(* Logix 5000 project; controller R400_500_XLS vendor 1 type 14 code 216 rev 31.11; software revision 31.01; part 4 of 32 *)
(* tags used below, declared in another part *)
   Alarm : SINT;   // Wait 3 seconds
   bResetAllCycle : BOOL;
   ClearIndex : DINT;
   Condenser : INT;
   Cycles : UDT_CYCLE[11];
   FINAL_RINSE_MAX_NBR : INT;   // Maximum nimber of final rinse
   LowPressAlmSp : REAL;   // Pump pressure too low setpoint
   MaxTrtTempSp : REAL;
   PrintoutMSGTranslation : DINT;   // Grapcet for Printout Message Translation
   PrintoutMSGTranslationONS : INT;
   PURE_WATER_HEATING_TIME : DINT;   // Time before an alarm is thrown when the pure water tank is heating
   PWTnkTempAlmSp : REAL;   // Pure water tank temperature too high setpoint
   String : STRING[50];   // String
   SumpTempAlmSp : REAL;   // Sump temperature too high setpoint
   tHandshakeToggle : TIMER;
   Tmr : TIMER[107];
   bFactoryReset : BOOL;
   bFactoryResetCompleted : BOOL;
   BoilingValue : REAL;
   bONSFactoryReset : BOOL;
   bResetHardwareOptions : BOOL;
   bResetModulesConfiguration : BOOL;
   bResetSystemOptions : BOOL;
   Cfg_10_Modules : BOOL;   // Chassis is configured 10 slots
   Cfg_11_Modules : BOOL;
   ChangeLanguage : BOOL;   // Tag Changed By HMI To Start Printout Message Translation
   COOLING_PHASE_TIME : DINT;   // Time of the cooling phase when time based drying
   CycleCounter : DINT;
   DrainExtensionTime : DINT;
   EmailSMSInt : INT[8];   // Email & SMS Notification Integer
   FC45_NbCycBeforeMaint : DINT;
   I_Chem_Cond : DINT;   // Chemical water conductivity
   I_Chm_1_Lvl_Sw : BOOL;   // Chemical Pump #1 level switch
   I_Chm_2_Lvl_Sw : BOOL;   // Chemical Pump #2 level switch
   I_Chm_3_Lvl_Sw : BOOL;   // Chemical Pump #3 level switch
   I_Chm_4_Lvl_Sw : BOOL;   // Chemical Pump #4 level switch
   I_Dry_RTD : DINT;   // Drying RTD
   I_Final_Rinse_Cond : DINT;   // Final rinse water conductivity
   I_Ld_Dr_Cls_Sw : BOOL;   // Load door close
   I_Ld_Dr_Obs_Sw : BOOL;   // Load door obstruction switch
   I_MCR : BOOL;   // MCR input
   I_Mtr_Ovrld : BOOL;   // Motor overload
   I_Pump_Press : DINT;   // Recirculation pump pressure
   I_Pure_Water_Filling_Auth : BOOL;
   I_Pw_Tnk_Lvl_Sw : BOOL;   // Pure water tank level switch
   I_Pw_Tnk_RTD : DINT;   // Pure water tank RTD
   I_Pw_Tnk_Sft_Lvl_Sw : BOOL;   // Pure water tank safety level switch
   I_Shlf_Sw : BOOL;   // Shelf switch
   I_Smp_Lvl_Hgh : BOOL;   // Sump high level switch
   I_Smp_Lvl_Lw : BOOL;   // Sump low level switch
   I_Smp_RTD : DINT;   // Sump RTD
   I_Smp_Sft_Lvl_Sw : BOOL;   // Sump safety level switch
   I_Unld_Dr_Cls_Sw : BOOL;   // Unload door close
   I_Unld_Dr_Obs_Sw : BOOL;   // Unload door obstruction switch
   I_UnldDr_ClseSlnce_Bttn : BOOL;   // Door Close/ Silence button Unload Side
   I_UnldDr_Opn_Bttn : BOOL;   // Door Open button Unload side
   iDelayBeforeFillingAuthAlarmMM : DINT;
   iDelayBeforeFillingAuthAlarmSS : DINT;
   iInactivityLogoutTime : DINT;   // Inactivity Logout Time In Minutes
   iPWClosingDelayMM : DINT;
   iPWClosingDelaySS : DINT;
   msg : BOOL[512];
   MsgIterator : DINT;   // Iterator to Iterate Through all Printout Mesage
   MsgNumbers : DINT;
   NOT_USED : SINT[3];
   NumInput : UDT_NUMERIC_INPUT[65];   // Numeric input
   NumInputReal : UDT_NUMERIC_INPUT_REAL[17];
   PrintoutMsgHandshake : BOOL;   // Flag Send to HMI to Acknowledge Reception of Message
   PrintoutMsgNotification : BOOL[512];   // Flag Send by HMI when a Message is sended to PLC
   Screen_Ctrl : DINT;   // PLC Screen Request
   SumpAlarmFillTime : DINT;
   Tpb : DINT[11];
   Unit : Hrdwre;   // Unit Configuration
(* MainProgram, continued *)

ROUTINE EMAIL_SEND   (* ladder *)
// SEND EMAIL
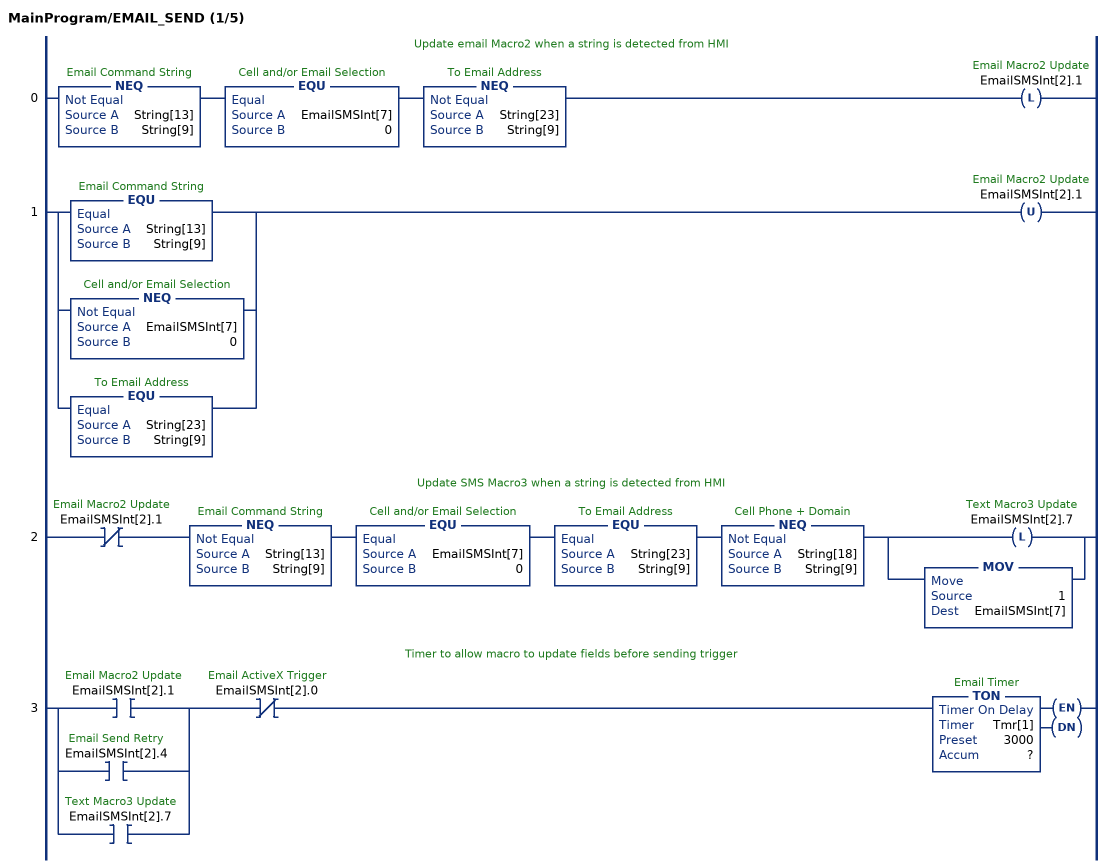
   // Update email Macro2 when a string is detected from HMI
   0: NEQ(String[13],String[9])EQU(EmailSMSInt[7],0)NEQ(String[23],String[9])OTL(EmailSMSInt[2].1);
   1: [EQU(String[13],String[9]) ,NEQ(EmailSMSInt[7],0) ,EQU(String[23],String[9]) ]OTU(EmailSMSInt[2].1);
   // Update SMS Macro3 when a string is detected from HMI
   2: XIO(EmailSMSInt[2].1)NEQ(String[13],String[9])EQU(EmailSMSInt[7],0)EQU(String[23],String[9])NEQ(String[18],String[9])[OTL(EmailSMSInt[2].7) ,MOV(1,EmailSMSInt[7]) ];
   // Timer to allow macro to update fields before sending trigger
   3: [XIC(EmailSMSInt[2].1) ,XIC(EmailSMSInt[2].4) ,XIC(EmailSMSInt[2].7) ]XIO(EmailSMSInt[2].0)TON(Tmr[1],?,?);
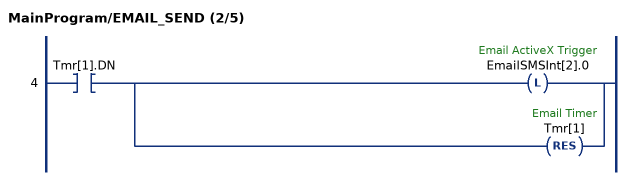
   4: XIC(Tmr[1].DN)[OTL(EmailSMSInt[2].0) ,RES(Tmr[1]) ];
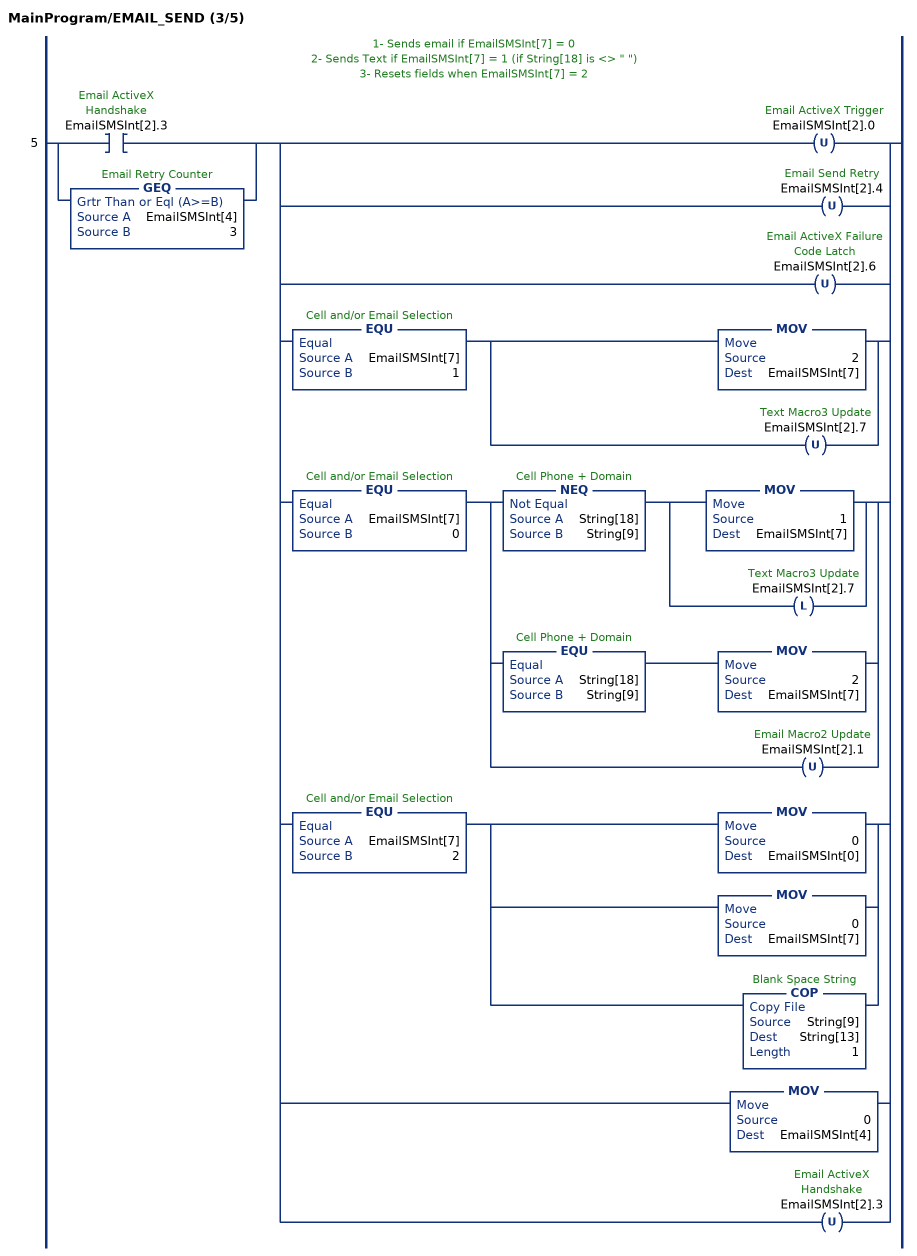
   // 1- Sends email if EmailSMSInt[7] = 0
   // 2- Sends Text if EmailSMSInt[7] = 1 (if String[18] is <> " ")
   // 3- Resets fields when EmailSMSInt[7] = 2
   5: [XIC(EmailSMSInt[2].3) ,GEQ(EmailSMSInt[4],3) ][OTU(EmailSMSInt[2].0) ,OTU(EmailSMSInt[2].4) ,OTU(EmailSMSInt[2].6) ,EQU(EmailSMSInt[7],1) [MOV(2,EmailSMSInt[7]) ,OTU(EmailSMSInt[2].7) ] ,EQU(EmailSMSInt[7],0) [NEQ(String[18],String[9]) [MOV(1,EmailSMSInt[7]) ,OTL(EmailSMSInt[2].7) ] ,EQU(String[18],String[9]) MOV(2,EmailSMSInt[7]) ,OTU(EmailSMSInt[2].1) ] ,EQU(EmailSMSInt[7],2) [MOV(0,EmailSMSInt[0]) ,MOV(0,EmailSMSInt[7]) ,COP(String[9],String[13],1) ] ,MOV(0,EmailSMSInt[4]) ,OTU(EmailSMSInt[2].3) ];
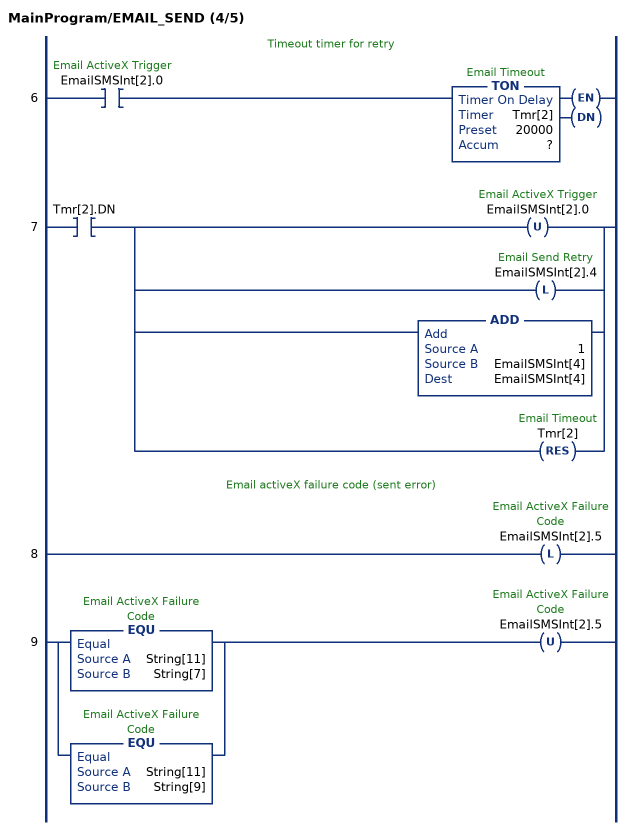
   // Timeout timer for retry
   6: XIC(EmailSMSInt[2].0)TON(Tmr[2],?,?);
   7: XIC(Tmr[2].DN)[OTU(EmailSMSInt[2].0) ,OTL(EmailSMSInt[2].4) ,ADD(1,EmailSMSInt[4],EmailSMSInt[4]) ,RES(Tmr[2]) ];
   // Email activeX failure code (sent error)
   8: OTL(EmailSMSInt[2].5);
   9: [EQU(String[11],String[7]) ,EQU(String[11],String[9]) ]OTU(EmailSMSInt[2].5);
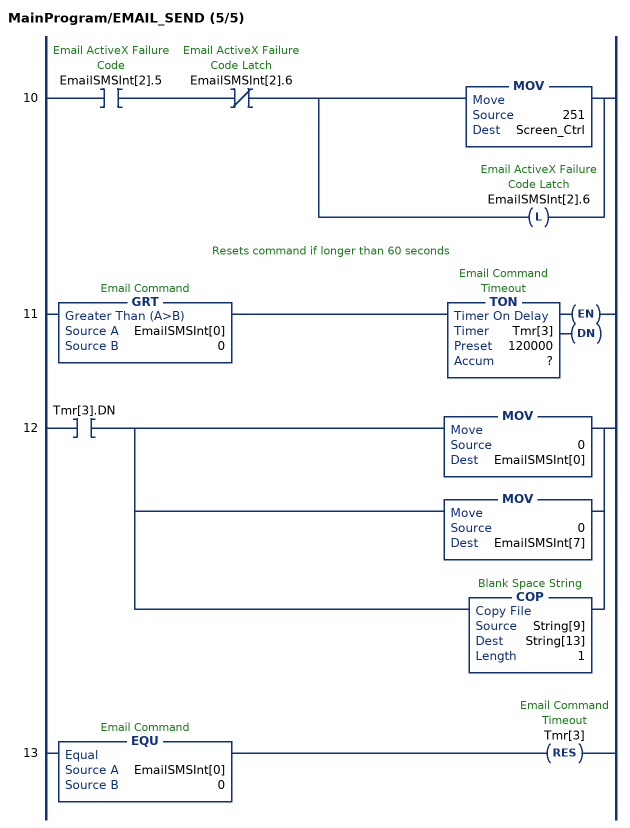
   10: XIC(EmailSMSInt[2].5)XIO(EmailSMSInt[2].6)[MOV(251,Screen_Ctrl) ,OTL(EmailSMSInt[2].6) ];
   // Resets command if longer than 60 seconds
   11: GRT(EmailSMSInt[0],0)TON(Tmr[3],?,?);
   12: XIC(Tmr[3].DN)[MOV(0,EmailSMSInt[0]) ,MOV(0,EmailSMSInt[7]) ,COP(String[9],String[13],1) ];
   13: EQU(EmailSMSInt[0],0)RES(Tmr[3]);
END_ROUTINE

ROUTINE FactoryReset   (* ladder *)
// This Routine contains logic to manage the Factory Reset
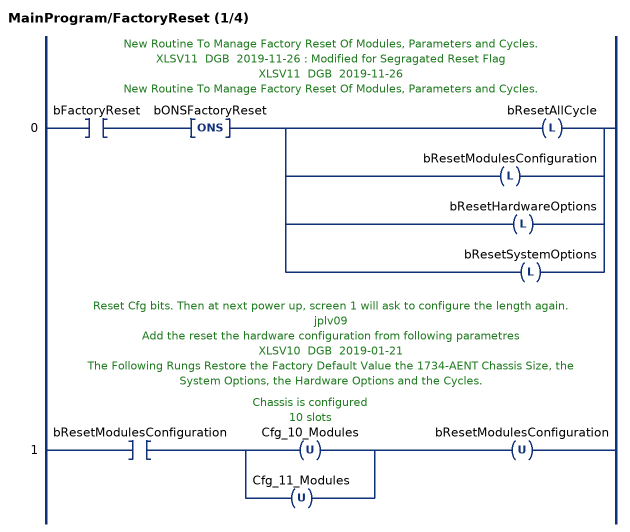
   // New Routine To Manage Factory Reset Of Modules, Parameters and Cycles.
   // XLSV11  DGB  2019-11-26 : Modified for Segragated Reset Flag
   // XLSV11  DGB  2019-11-26
   // New Routine To Manage Factory Reset Of Modules, Parameters and Cycles.
   0: XIC(bFactoryReset)ONS(bONSFactoryReset)[OTL(bResetAllCycle) ,OTL(bResetModulesConfiguration) ,OTL(bResetHardwareOptions) ,OTL(bResetSystemOptions) ];
   // Reset Cfg bits. Then at next power up, screen 1 will ask to configure the length again.
   // jplv09
   // Add the reset the hardware configuration from following parametres
   // XLSV10  DGB  2019-01-21
   // The Following Rungs Restore the Factory Default Value the 1734-AENT Chassis Size, the System Options, the Hardware Options and the Cycles.
   1: XIC(bResetModulesConfiguration)[OTU(Cfg_10_Modules) ,OTU(Cfg_11_Modules) ]OTU(bResetModulesConfiguration);
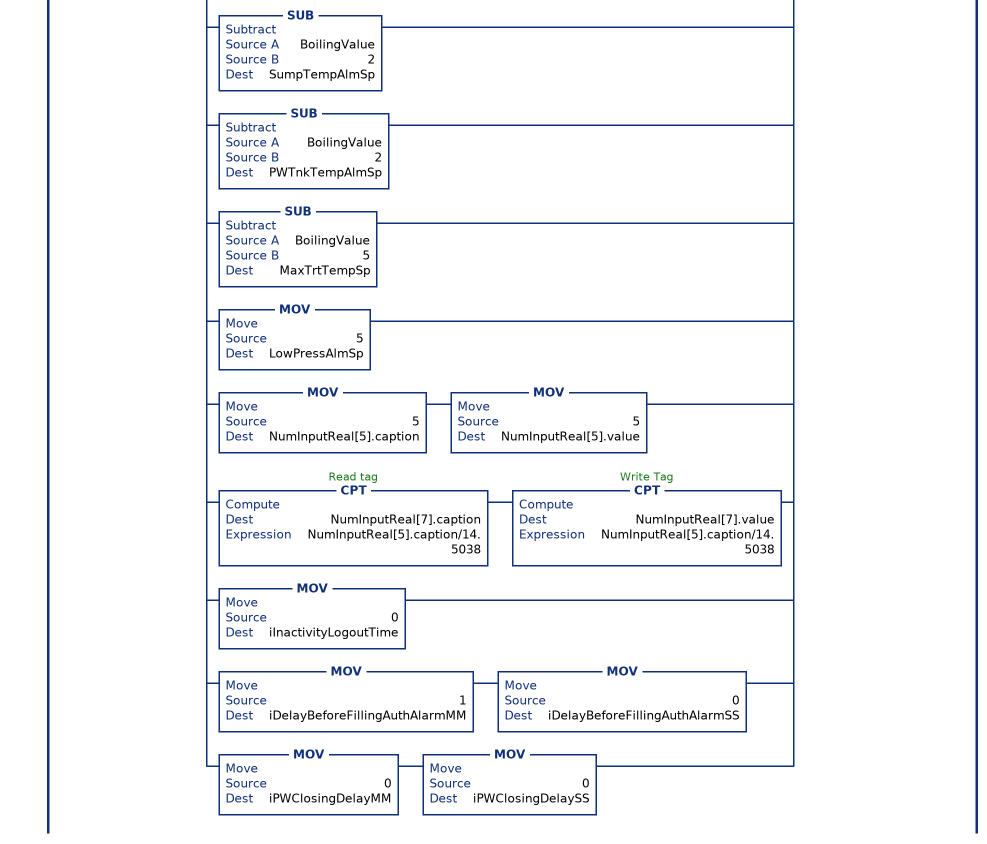
   // XLSV10  DGB  2019-01-21
   // New Rung to Restore the Factory Default Value of System Options
   // XLSV13  DGB  2021-03-16 : PW Filling Handshake : Added Pure Water Closing Delay & Delay Before Fill Auth Alarm Message
   2: XIC(bResetSystemOptions)[MOV(0,CycleCounter) ,MOV(1000,FC45_NbCycBeforeMaint) ,[MOV(120000,SumpAlarmFillTime) ,MOV(2,NumInput[9].caption) MOV(2,NumInput[9].value) ,MOV(0,NumInput[10].caption) MOV(0,NumInput[10].value) ] ,[MOV(20000,Tmr[88].PRE) ,MOV(20,NumInput[52].caption) MOV(20,NumInput[52].value) ] ,[MOV(480000,Tmr[37].PRE) ,MOV(8,NumInput[38].caption) MOV(8,NumInput[38].value) ,MOV(0,NumInput[39].caption) MOV(0,NumInput[39].value) ] ,[MOV(1200000,PURE_WATER_HEATING_TIME) ,MOV(20,NumInput[40].caption) MOV(20,NumInput[40].value) ,MOV(0,NumInput[41].caption) MOV(0,NumInput[41].value) ] ,[MOV(9,FINAL_RINSE_MAX_NBR) ,MOV(9,NumInput[42].caption) MOV(9,NumInput[42].value) ] ,[MOV(0,DrainExtensionTime) ,MOV(0,NumInput[43].caption) MOV(0,NumInput[43].value) ] ,[MOV(120000,Tmr[31].PRE) ,MOV(2,NumInput[44].caption) MOV(2,NumInput[44].value) ,MOV(0,NumInput[45].caption) MOV(0,NumInput[45].value) ] ,[MOV(120000,COOLING_PHASE_TIME) ,MOV(2,NumInput[47].caption) MOV(2,NumInput[47].value) ,MOV(0,NumInput[48].caption) MOV(0,NumInput[48].value) ] ,[MOV(0,NumInput[46].caption) MOV(0,NumInput[46].value) ,CPT(BoilingValue,100.03) ,SUB(BoilingValue,2,SumpTempAlmSp) ,SUB(BoilingValue,2,PWTnkTempAlmSp) ,SUB(BoilingValue,5,MaxTrtTempSp) ] ,[MOV(5,LowPressAlmSp) ,MOV(5,NumInputReal[5].caption) MOV(5,NumInputReal[5].value) ,CPT(NumInputReal[7].caption,NumInputReal[5].caption/14.5038) CPT(NumInputReal[7].value,NumInputReal[5].caption/14.5038) ] ,MOV(0,iInactivityLogoutTime) ,MOV(1,iDelayBeforeFillingAuthAlarmMM) MOV(0,iDelayBeforeFillingAuthAlarmSS) ,MOV(0,iPWClosingDelayMM) MOV(0,iPWClosingDelaySS) ]OTU(bResetSystemOptions);
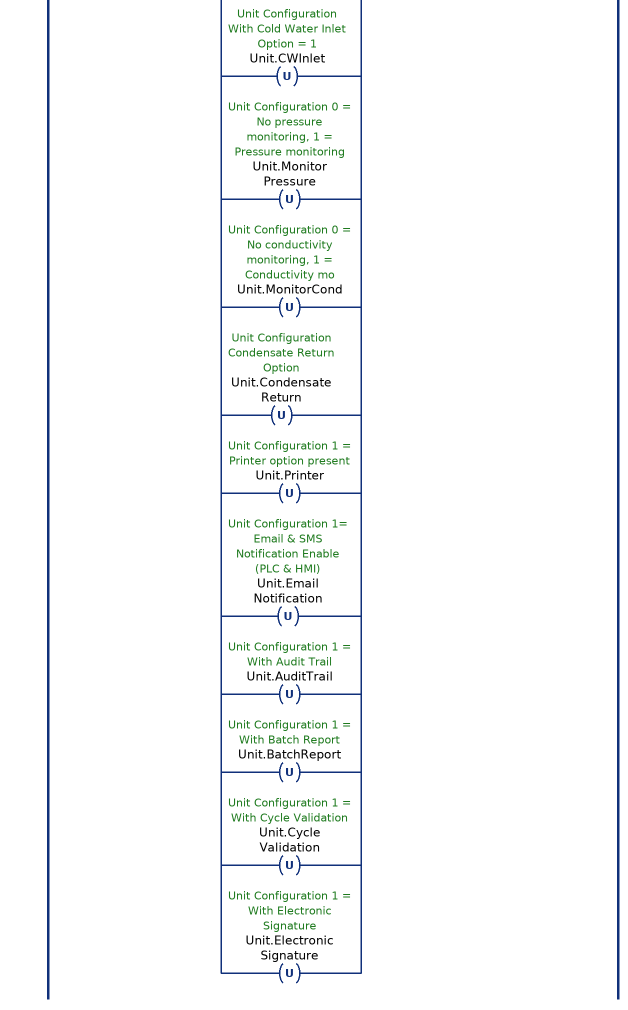
   // XLSV10  DGB  2019-01-21
   // New Rung to Restore the Factory Default Value of Hardware Options
   // XLSV11 DGB 2019-11-26
   // Modified To Latch Batch Report & Audit Trail
   // XLSV13  DGB  2021-04-01 : Cycle Validation & Electronic Signature
   3: XIC(bResetHardwareOptions)[OTU(Unit.Model) ,OTU(Unit.NbDoors) ,OTU(Unit.PreWtrTnk) ,OTU(Unit.HtRcvryTnk) ,[OTU(Unit.Dry) ,OTU(Tpb[7].10) ,OTU(Tpb[7].11) ,OTU(Tpb[7].12) ] ,OTU(Unit.ElectricUnit) ,OTU(Unit.CoolDown) ,OTU(Tpb[7].13) ,OTU(Unit.Condenser) ,OTU(Unit.CWInlet) ,OTU(Unit.MonitorPressure) ,OTU(Unit.MonitorCond) ,OTU(Unit.CondensateReturn) ,OTU(Unit.Printer) ,OTU(Unit.EmailNotification) ,OTU(Unit.AuditTrail) ,OTU(Unit.BatchReport) ,OTU(Unit.CycleValidation) ,OTU(Unit.ElectronicSignature) ]OTU(bResetHardwareOptions);
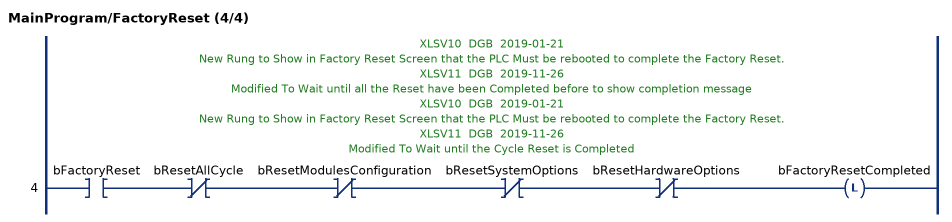
   // XLSV10  DGB  2019-01-21
   // New Rung to Show in Factory Reset Screen that the PLC Must be rebooted to complete the Factory Reset.
   // XLSV11  DGB  2019-11-26
   // Modified To Wait until all the Reset have been Completed before to show completion message
   // XLSV10  DGB  2019-01-21
   // New Rung to Show in Factory Reset Screen that the PLC Must be rebooted to complete the Factory Reset.
   // XLSV11  DGB  2019-11-26
   // Modified To Wait until the Cycle Reset is Completed
   4: XIC(bFactoryReset)XIO(bResetAllCycle)XIO(bResetModulesConfiguration)XIO(bResetSystemOptions)XIO(bResetHardwareOptions)OTL(bFactoryResetCompleted);
END_ROUTINE

ROUTINE HandshakeToTransMSG   (* ladder *)
// The message send from the HMI to PLC request a Handshake.
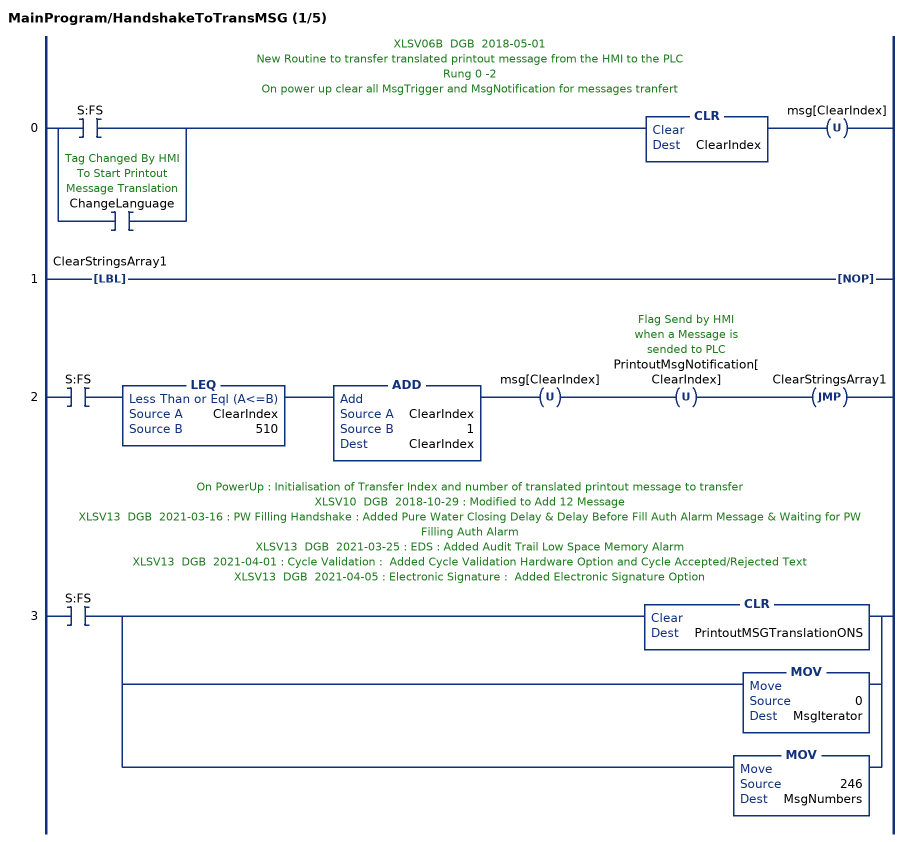
   // XLSV06B  DGB  2018-05-01
   //  New Routine to transfer translated printout message from the HMI to the PLC
   // Rung 0 -2
   // On power up clear all MsgTrigger and MsgNotification for messages tranfert
   0: [XIC(S:FS) ,XIC(ChangeLanguage) ]CLR(ClearIndex)OTU(msg[ClearIndex]);
   1: LBL(ClearStringsArray1)NOP();
   2: XIC(S:FS)LEQ(ClearIndex,510)ADD(ClearIndex,1,ClearIndex)OTU(msg[ClearIndex])OTU(PrintoutMsgNotification[ClearIndex])JMP(ClearStringsArray1);
   // On PowerUp : Initialisation of Transfer Index and number of translated printout message to transfer
   // XLSV10  DGB  2018-10-29 : Modified to Add 12 Message
   // XLSV13  DGB  2021-03-16 : PW Filling Handshake : Added Pure Water Closing Delay & Delay Before Fill Auth Alarm Message & Waiting for PW Filling Auth Alarm
   // XLSV13  DGB  2021-03-25 : EDS : Added Audit Trail Low Space Memory Alarm
   // XLSV13  DGB  2021-04-01 : Cycle Validation :  Added Cycle Validation Hardware Option and Cycle Accepted/Rejected Text
   // XLSV13  DGB  2021-04-05 : Electronic Signature :  Added Electronic Signature Option
   3: XIC(S:FS)[CLR(PrintoutMSGTranslationONS) ,MOV(0,MsgIterator) ,MOV(246,MsgNumbers) ];
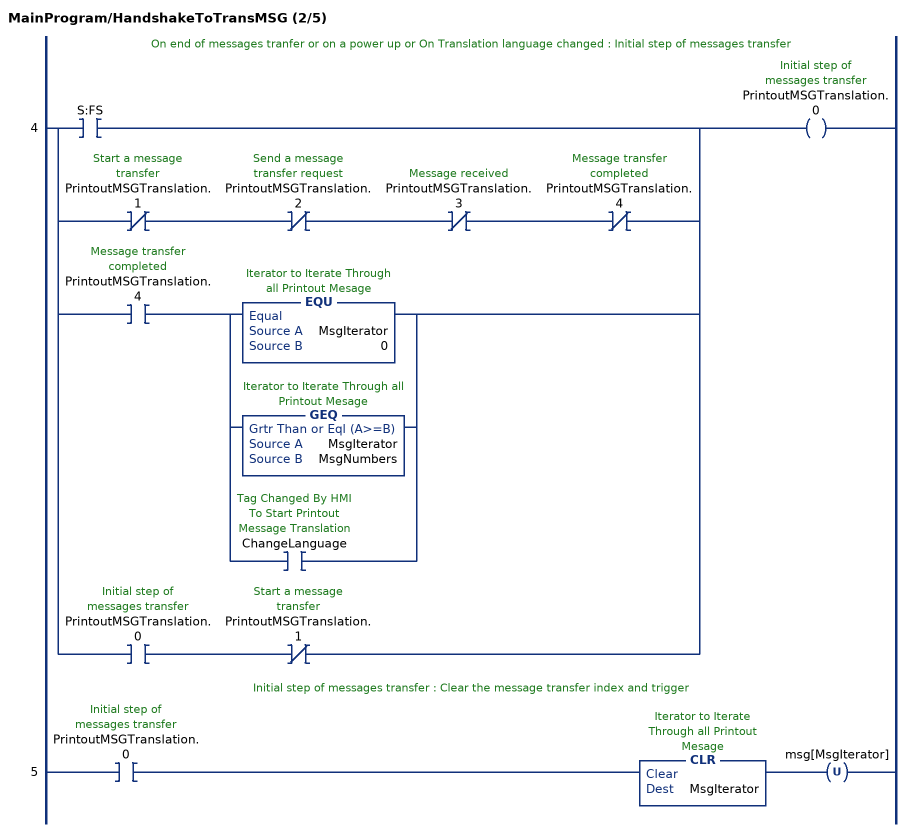
   // On end of messages tranfer or on a power up or On Translation language changed : Initial step of messages transfer
   4: [XIC(S:FS) ,XIO(PrintoutMSGTranslation.1) XIO(PrintoutMSGTranslation.2) XIO(PrintoutMSGTranslation.3) XIO(PrintoutMSGTranslation.4) ,XIC(PrintoutMSGTranslation.4) [EQU(MsgIterator,0) ,GEQ(MsgIterator,MsgNumbers) ,XIC(ChangeLanguage) ] ,XIC(PrintoutMSGTranslation.0) XIO(PrintoutMSGTranslation.1) ]OTE(PrintoutMSGTranslation.0);
   // Initial step of messages transfer : Clear the message transfer index and trigger
   5: XIC(PrintoutMSGTranslation.0)CLR(MsgIterator)OTU(msg[MsgIterator]);
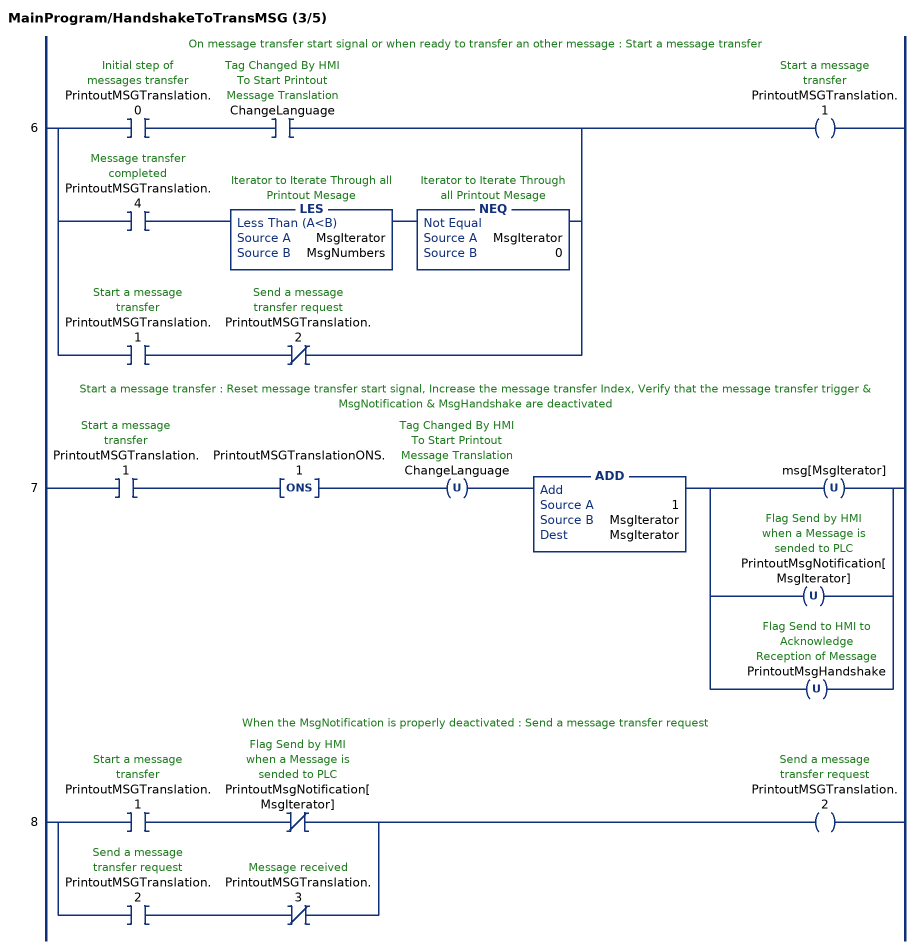
   // On message transfer start signal or when ready to transfer an other message : Start a message transfer
   6: [XIC(PrintoutMSGTranslation.0) XIC(ChangeLanguage) ,XIC(PrintoutMSGTranslation.4) LES(MsgIterator,MsgNumbers) NEQ(MsgIterator,0) ,XIC(PrintoutMSGTranslation.1) XIO(PrintoutMSGTranslation.2) ]OTE(PrintoutMSGTranslation.1);
   // Start a message transfer : Reset message transfer start signal, Increase the message transfer Index, Verify that the message transfer trigger & MsgNotification & MsgHandshake are deactivated
   7: XIC(PrintoutMSGTranslation.1)ONS(PrintoutMSGTranslationONS.1)OTU(ChangeLanguage)ADD(1,MsgIterator,MsgIterator)[OTU(msg[MsgIterator]) ,OTU(PrintoutMsgNotification[MsgIterator]) ,OTU(PrintoutMsgHandshake) ];
   // When the MsgNotification is properly deactivated : Send a message transfer request
   8: [XIC(PrintoutMSGTranslation.1) XIO(PrintoutMsgNotification[MsgIterator]) ,XIC(PrintoutMSGTranslation.2) XIO(PrintoutMSGTranslation.3) ]OTE(PrintoutMSGTranslation.2);
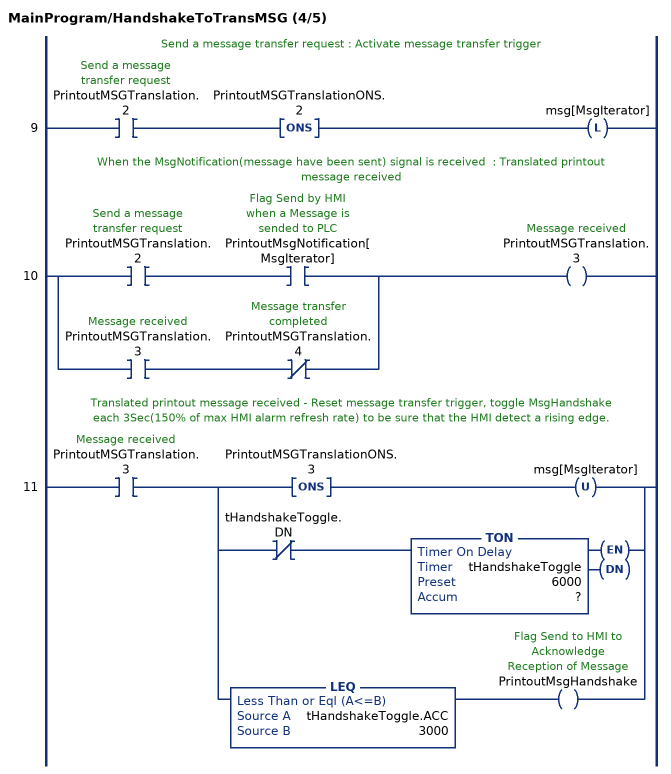
   // Send a message transfer request : Activate message transfer trigger
   9: XIC(PrintoutMSGTranslation.2)ONS(PrintoutMSGTranslationONS.2)OTL(msg[MsgIterator]);
   // When the MsgNotification(message have been sent) signal is received  : Translated printout message received
   10: [XIC(PrintoutMSGTranslation.2) XIC(PrintoutMsgNotification[MsgIterator]) ,XIC(PrintoutMSGTranslation.3) XIO(PrintoutMSGTranslation.4) ]OTE(PrintoutMSGTranslation.3);
   // Translated printout message received - Reset message transfer trigger, toggle MsgHandshake each 3Sec(150% of max HMI alarm refresh rate) to be sure that the HMI detect a rising edge.
   11: XIC(PrintoutMSGTranslation.3)[ONS(PrintoutMSGTranslationONS.3) OTU(msg[MsgIterator]) ,XIO(tHandshakeToggle.DN) TON(tHandshakeToggle,?,?) ,LEQ(tHandshakeToggle.ACC,3000) OTE(PrintoutMsgHandshake) ];
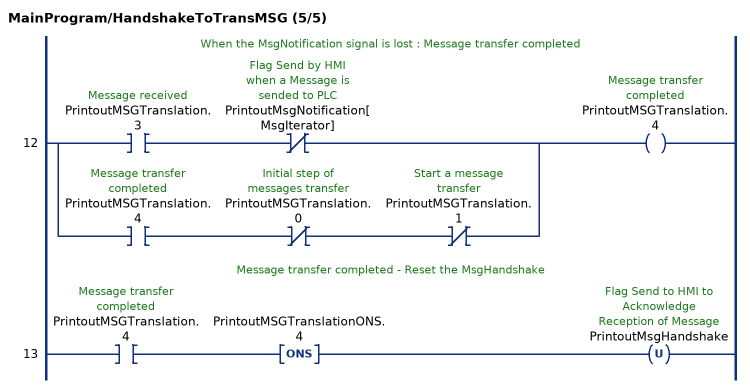
   // When the MsgNotification signal is lost : Message transfer completed
   12: [XIC(PrintoutMSGTranslation.3) XIO(PrintoutMsgNotification[MsgIterator]) ,XIC(PrintoutMSGTranslation.4) XIO(PrintoutMSGTranslation.0) XIO(PrintoutMSGTranslation.1) ]OTE(PrintoutMSGTranslation.4);
   // Message transfer completed - Reset the MsgHandshake
   13: XIC(PrintoutMSGTranslation.4)ONS(PrintoutMSGTranslationONS.4)OTU(PrintoutMsgHandshake);
END_ROUTINE

ROUTINE Inputs   (* ladder *)
// The routine maps the point i/o inputs
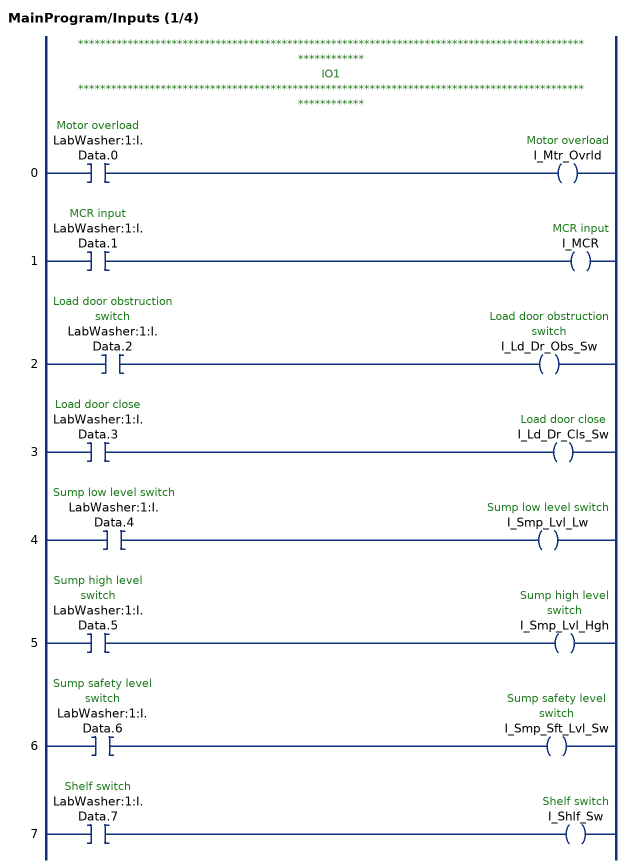
   // ********************************************************************************************************
   // IO1
   // ********************************************************************************************************
   0: XIC(LabWasher:1:I.Data.0)OTE(I_Mtr_Ovrld);
   1: XIC(LabWasher:1:I.Data.1)OTE(I_MCR);
   2: XIC(LabWasher:1:I.Data.2)OTE(I_Ld_Dr_Obs_Sw);
   3: XIC(LabWasher:1:I.Data.3)OTE(I_Ld_Dr_Cls_Sw);
   4: XIC(LabWasher:1:I.Data.4)OTE(I_Smp_Lvl_Lw);
   5: XIC(LabWasher:1:I.Data.5)OTE(I_Smp_Lvl_Hgh);
   6: XIC(LabWasher:1:I.Data.6)OTE(I_Smp_Sft_Lvl_Sw);
   7: XIC(LabWasher:1:I.Data.7)OTE(I_Shlf_Sw);
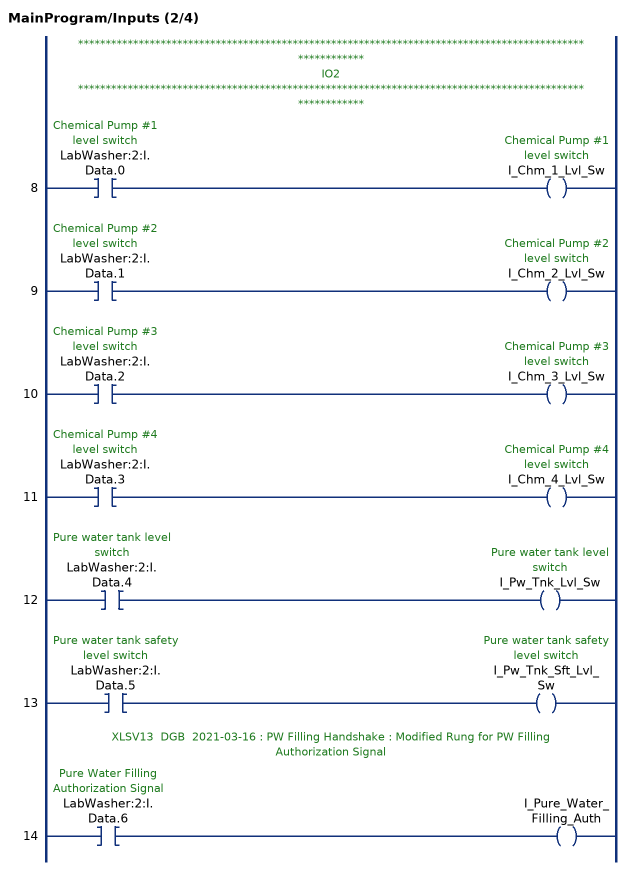
   // ********************************************************************************************************
   // IO2
   // ********************************************************************************************************
   8: XIC(LabWasher:2:I.Data.0)OTE(I_Chm_1_Lvl_Sw);
   9: XIC(LabWasher:2:I.Data.1)OTE(I_Chm_2_Lvl_Sw);
   10: XIC(LabWasher:2:I.Data.2)OTE(I_Chm_3_Lvl_Sw);
   11: XIC(LabWasher:2:I.Data.3)OTE(I_Chm_4_Lvl_Sw);
   12: XIC(LabWasher:2:I.Data.4)OTE(I_Pw_Tnk_Lvl_Sw);
   13: XIC(LabWasher:2:I.Data.5)OTE(I_Pw_Tnk_Sft_Lvl_Sw);
   // XLSV13  DGB  2021-03-16 : PW Filling Handshake : Modified Rung for PW Filling Authorization Signal
   14: XIC(LabWasher:2:I.Data.6)OTE(I_Pure_Water_Filling_Auth);
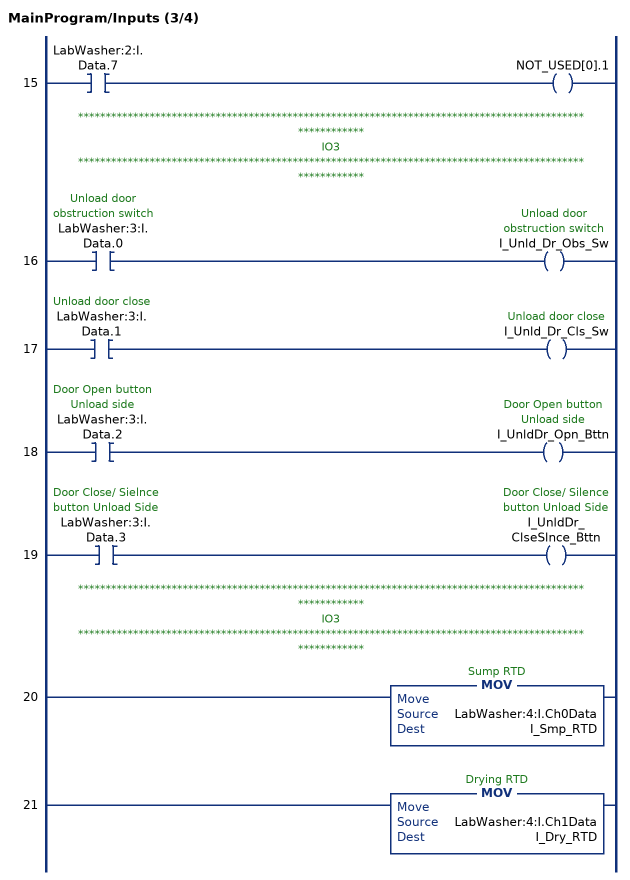
   15: XIC(LabWasher:2:I.Data.7)OTE(NOT_USED[0].1);
   // ********************************************************************************************************
   // IO3
   // ********************************************************************************************************
   16: XIC(LabWasher:3:I.Data.0)OTE(I_Unld_Dr_Obs_Sw);
   17: XIC(LabWasher:3:I.Data.1)OTE(I_Unld_Dr_Cls_Sw);
   18: XIC(LabWasher:3:I.Data.2)OTE(I_UnldDr_Opn_Bttn);
   19: XIC(LabWasher:3:I.Data.3)OTE(I_UnldDr_ClseSlnce_Bttn);
   // ********************************************************************************************************
   // IO3
   // ********************************************************************************************************
   20: MOV(LabWasher:4:I.Ch0Data,I_Smp_RTD);
   21: MOV(LabWasher:4:I.Ch1Data,I_Dry_RTD);
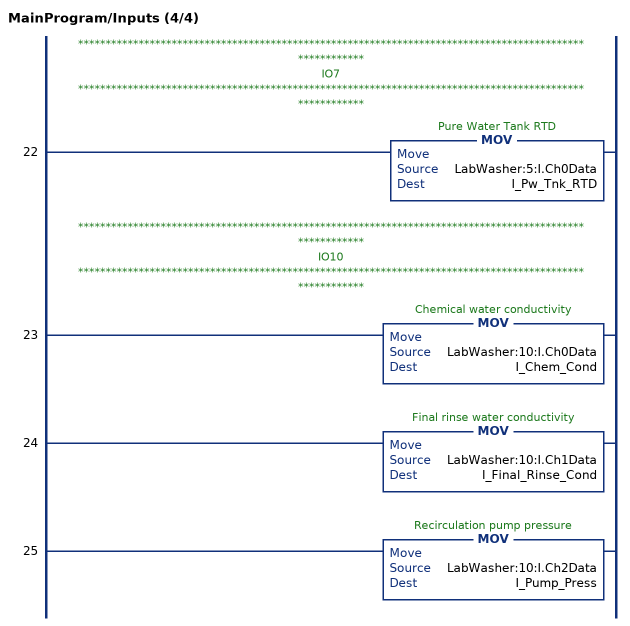
   // ********************************************************************************************************
   // IO7
   // ********************************************************************************************************
   22: MOV(LabWasher:5:I.Ch0Data,I_Pw_Tnk_RTD);
   // ********************************************************************************************************
   // IO10
   // ********************************************************************************************************
   23: MOV(LabWasher:10:I.Ch0Data,I_Chem_Cond);
   24: MOV(LabWasher:10:I.Ch1Data,I_Final_Rinse_Cond);
   25: MOV(LabWasher:10:I.Ch2Data,I_Pump_Press);
END_ROUTINE
